Fanuc KAREL source: kd00041.KL

-- PROVISIONAL review KL for V1013-1; original PC SHA256 90151307fc0de7ca67f5bfcd60f91c68007dfaf0f9090433d241f30662490399
-- Incomplete behavior may be omitted. Consult companion uncertainty JSON. Do not deploy.
PROGRAM KD00041
%NOLOCKGROUP
BEGIN
  -- UNRESOLVED_PC offsets 5-12; opcodes 9D,23
  -- UNRESOLVED_PC offsets 17-21; opcodes 7F
END KD00041
